// TIA Portal V21 export
Screen "R06c_MoveH"  1024x768, Number=46, Template=Tpl
  ScreenLayer 
    IOField "P_CraneX" at 10,10 size 100x30  Mode=Output
      ProcessValue := P_Cell
      HorizontalMovementAnimation "HorizontalMovementAnimation"
        tag P_Cell
